(* IEC 61131-3 sources: guidance-for-physical-ai-production-designer-on-aws/source/plan2cell/examples/cell_2robot/plc/codesys/robots/robot1/GVL, 3 files *)

(* ---- GVL_DeviceParams.st ---- *)
(*
 * GVL_DeviceParams
 * PROFINET device identity parameters.
 * Device simulator R1 (robot1, station kuka-robi1), cell cell_2robot. Generated by bt2plc 0.1.0.
 *
 * These parameters configure how the CODESYS PROFINET Device presents itself
 * on the network. They MUST match what the Siemens PLC expects (from the GSDML).
 *
 * In CODESYS, these are typically set via:
 *   1. The "PROFINET Device IEC Objects" tab in the device editor
 *   2. Or programmatically by writing to the device parameter structure
 *
 * The CODESYS PROFINET Device stack reads these at startup and uses them
 * in DCP responses and during the PROFINET connection establishment.
 *
 * IMPORTANT: The default CODESYS values (VendorId=0x02CC, DeviceId=0x1017)
 * will NOT work with the Siemens PLC that expects KUKA (0x019B / 0x0301).
 * You MUST override them.
 *)

{attribute 'qualified_only'}
VAR_GLOBAL CONSTANT
    (* === KUKA VKRCnexxt Device Identity === *)
    (* These values come from GSDML-V2.25-KUKA-Roboter-GmbH-VKR C4-Device-V1.0 *)

    VENDOR_ID           : UINT        := 16#019B;                 (* KUKA Roboter GmbH *)
    DEVICE_ID           : UINT        := 16#0301;                 (* VKR C4 Device *)
    STATION_TYPE        : STRING(240) := 'KUKA VKR C4';           (* Station type string *)
    DEVICE_TYPE         : STRING(28)  := 'KUKA VKR C4';           (* Device type string *)
    ORDER_ID            : STRING(20)  := 'KUKA VKRC nexxt';       (* Order number *)
    HW_REVISION         : UINT        := 1;                       (* Hardware revision *)
    SW_REV_PREFIX       : USINT       := 16#56;                   (* 'V' in ASCII *)
    SW_REV_MAJOR        : UINT        := 8;                       (* V8.x *)
    SW_REV_MINOR        : UINT        := 2;                       (* x.2 *)
    SW_REV_PATCH        : UINT        := 0;                       (* x.x.0 *)

    (* === Module Identification Numbers (from GSDML) === *)
    MODULE_IDENT_DAP    : DWORD       := DWORD#16#00000301;       (* DAP - Slot 0 *)
    MODULE_IDENT_FDIO64 : DWORD       := DWORD#16#0000008F;       (* PROFIsafe - Slot 1 *)
    MODULE_IDENT_DIO256 : DWORD       := DWORD#16#00001000;       (* VASS telegram - Slot 2 *)
    SUBMODULE_IDENT     : DWORD       := DWORD#16#00000001;       (* Submodule ident (all slots) *)

    (* === PROFIsafe Parameters (Slot 1) === *)
    (* These must match the F-parameter record in the PLC safety configuration *)
    F_SIL_LEVEL         : UINT        := 3;                       (* SIL 3 *)
    F_CRC_LENGTH        : UINT        := 3;                       (* 3-byte CRC *)
    F_WD_TIME_DEFAULT   : UINT        := 500;                     (* Watchdog 500ms *)
    F_BLOCK_ID          : UINT        := 0;                       (* Block ID *)
    F_PAR_CRC_DEFAULT   : UINT        := 16#FF59;                 (* Default F_Par_CRC = 65369 *)
END_VAR

(* ---- GVL_IO.st ---- *)
(*
 * GVL_IO
 * Global variable list for the PROFINET device I/O mapping.
 * Device simulator R1 (robot1, station kuka-robi1), cell cell_2robot. Generated by bt2plc 0.1.0.
 *
 * These variables are mapped to the PROFINET device modules via the I/O Mapping tab.
 * Do NOT use AT addresses - the mapping is done in the device configuration.
 * Only PLC_PRG accesses this GVL: it copies the commands into local images and writes
 * the robot status back as a whole array / as scalars (the FBs never touch GVL_IO).
 *
 * Module mapping (set in I/O Mapping tab of each module):
 *   SafeIO_FDIO64 (Slot 1):
 *     "8 safe digital inputs" channels  -> GVL_IO.bySafeIn0..bySafeIn7
 *     "8 safe digital outputs" channels -> GVL_IO.bySafeOut0..bySafeOut7
 *
 *   VASS_DIO256 (Slot 2):
 *     Input channel  -> GVL_IO.aVassInputData
 *     Output channel -> GVL_IO.aVassOutputData
 *)

{attribute 'qualified_only'}
VAR_GLOBAL
    (* ========================================================================
       SLOT 1 - PROFIsafe FDIO64 Module
       8 individual USINT/BYTE channels per direction
       Map each one to the corresponding "8 safe digital inputs/outputs" row
       ======================================================================== *)

    (* Safe Inputs: Robot -> PLC (mapped to "8 safe digital inputs" channels) *)
    bySafeIn0       : BYTE;     (* Safe input byte 0: Drive status *)
    bySafeIn1       : BYTE;     (* Safe input byte 1: Gate/protection *)
    bySafeIn2       : BYTE;     (* Safe input byte 2: STO/SS1/SS2/SOS/SLS *)
    bySafeIn3       : BYTE;     (* Safe input byte 3: User *)
    bySafeIn4       : BYTE;     (* Safe input byte 4: User *)
    bySafeIn5       : BYTE;     (* Safe input byte 5: User *)
    bySafeIn6       : BYTE;     (* Safe input byte 6: User *)
    bySafeIn7       : BYTE;     (* Safe input byte 7: User *)

    (* Safe Outputs: PLC -> Robot (mapped to "8 safe digital outputs" channels) *)
    bySafeOut0      : BYTE;     (* Safe output byte 0: Drive enable, E-Stop, SS1/SS2 *)
    bySafeOut1      : BYTE;     (* Safe output byte 1: Zone enables *)
    bySafeOut2      : BYTE;     (* Safe output byte 2: User *)
    bySafeOut3      : BYTE;     (* Safe output byte 3: User *)
    bySafeOut4      : BYTE;     (* Safe output byte 4: User *)
    bySafeOut5      : BYTE;     (* Safe output byte 5: User *)
    bySafeOut6      : BYTE;     (* Safe output byte 6: User *)
    bySafeOut7      : BYTE;     (* Safe output byte 7: User *)

    (* ========================================================================
       SLOT 2 - DIO256 VASS Telegram
       32 bytes per direction as arrays
       ======================================================================== *)

    (* VASS Inputs: Robot -> PLC (32 bytes) *)
    aVassInputData      : ARRAY[0..31] OF BYTE;

    (* VASS Outputs: PLC -> Robot (32 bytes) *)
    aVassOutputData     : ARRAY[0..31] OF BYTE;
END_VAR

(* ---- GVL_Program.st ---- *)
(*
 * GVL_Program - generated by bt2plc 0.1.0 - DO NOT EDIT
 * Robot program of robot1 (R1) for plan bt_1791274820_cell_2robot (cell cell_2robot)
 * Angles in degrees (KUKA A1..A6 after joint sign/offset), times in seconds from op start.
 *)
{attribute 'qualified_only'}
VAR_GLOBAL CONSTANT
    (* ========================================================================
       IDENTITY / PROTOCOL
       ======================================================================== *)
    ROBOT_TAG               : STRING(16) := 'R1';
    ROBOT_NS                : STRING(32) := 'robot1';
    ROBOT_INDEX             : WORD := WORD#1;
    PLAN_ID                 : WORD := WORD#16#A312;             (* must match the head PLC *)
    PROD_FOLGE              : WORD := WORD#11;
    HOME_FOLGE              : WORD := WORD#125;
    JOB_NUMBER_BYTE         : BOOL := FALSE;
    STEP_BYTE               : INT := 4;
    REQ_BYTE                : INT := 28;
    GRANT_BYTE              : INT := 12;
    PLAN_ID_BYTE            : INT := 4;
    R_TASK_S                : REAL := 0.0200;                   (* device MainTask interval *)
    R_HOME_S                : REAL := 7.0000;                   (* blind home duration *)
    R_AT_HOME_TOL_DEG       : REAL := 0.5000;
    R_START_TOL_DEG         : REAL := 1.0000;
    ERR_UNKNOWN_FOLGE       : WORD := WORD#16#0101;
    ERR_PLAN_MISMATCH       : WORD := WORD#16#0103;
    WARN_START_DEVIATION    : WORD := WORD#16#0201;

    (* ========================================================================
       PROGRAM
       ======================================================================== *)
    N_OPS                   : INT := 2;
    N_WP                    : INT := 27;
    arHomeDeg               : ARRAY[1..6] OF REAL := [0.0000, -90.0000, 90.0000, 0.0000, 0.0000, 0.0000];
    aOps                    : ARRAY[1..2] OF ST_OpDef := [
        (sName := 'STAGE_R1', nFirstWp := 1, nLastWp := 14, dwZoneMask := DWORD#16#00000000, tDelay := T#0MS, tHold := T#500MS, rDelay_s := 0.0000, rHold_s := 0.5000, rVelScale := 1.0000, bBlindHome := FALSE),    (* #1 STAGE_R1 (move) *)
        (sName := 'HOME', nFirstWp := 15, nLastWp := 27, dwZoneMask := DWORD#16#00000000, tDelay := T#0MS, tHold := T#0MS, rDelay_s := 0.0000, rHold_s := 0.0000, rVelScale := 1.0000, bBlindHome := FALSE)    (* #2 HOME (home) *)
    ];
    aWp                     : ARRAY[1..27] OF ST_Waypoint := [
        (* op 1 STAGE_R1 - traj_robot1_STAGE_R1 *)
        (rT := 0.0000, rA1 := 0.0000, rA2 := -90.0000, rA3 := 90.0000, rA4 := 0.0000, rA5 := 0.0000, rA6 := 0.0000),
        (rT := 0.2767, rA1 := 0.1421, rA2 := -89.0006, rA3 := 89.9771, rA4 := 0.0000, rA5 := 0.0000, rA6 := 0.0000),
        (rT := 0.5530, rA1 := 0.5354, rA2 := -86.2310, rA3 := 89.9133, rA4 := 0.0000, rA5 := 0.0000, rA6 := 0.0000),
        (rT := 0.8297, rA1 := 1.1310, rA2 := -82.0342, rA3 := 89.8161, rA4 := 0.0000, rA5 := 0.0000, rA6 := 0.0000),
        (rT := 1.1063, rA1 := 1.8795, rA2 := -76.7531, rA3 := 89.6931, rA4 := 0.0000, rA5 := 0.0000, rA6 := 0.0000),
        (rT := 1.3830, rA1 := 2.7319, rA2 := -70.7305, rA3 := 89.5515, rA4 := 0.0000, rA5 := 0.0000, rA6 := 0.0000),
        (rT := 1.6593, rA1 := 3.6388, rA2 := -64.3095, rA3 := 89.3990, rA4 := 0.0000, rA5 := 0.0000, rA6 := 0.0000),
        (rT := 1.9360, rA1 := 4.5513, rA2 := -57.8329, rA3 := 89.2429, rA4 := 0.0000, rA5 := 0.0000, rA6 := 0.0000),
        (rT := 2.2127, rA1 := 5.4200, rA2 := -51.6436, rA3 := 89.0908, rA4 := 0.0000, rA5 := 0.0000, rA6 := 0.0000),
        (rT := 2.4893, rA1 := 6.1959, rA2 := -46.0847, rA3 := 88.9501, rA4 := 0.0000, rA5 := 0.0000, rA6 := 0.0000),
        (rT := 2.7657, rA1 := 6.8297, rA2 := -41.4990, rA3 := 88.8283, rA4 := 0.0000, rA5 := 0.0000, rA6 := 0.0000),
        (rT := 3.0423, rA1 := 7.2722, rA2 := -38.2294, rA3 := 88.7329, rA4 := 0.0000, rA5 := 0.0000, rA6 := 0.0000),
        (rT := 3.1357, rA1 := 7.7267, rA2 := -33.2119, rA3 := 88.3788, rA4 := 0.0000, rA5 := 0.0000, rA6 := 0.0000),
        (rT := 3.2287, rA1 := 7.2722, rA2 := -35.0616, rA3 := 88.2443, rA4 := 0.0000, rA5 := 0.0000, rA6 := 0.0000),
        (* op 2 HOME - traj_robot1_n3 *)
        (rT := 0.0000, rA1 := 7.2722, rA2 := -35.0616, rA3 := 88.2443, rA4 := 0.0000, rA5 := 0.0000, rA6 := 0.0000),
        (rT := 0.2015, rA1 := 7.1292, rA2 := -36.1426, rA3 := 88.2788, rA4 := 0.0000, rA5 := 0.0000, rA6 := 0.0000),
        (rT := 0.4032, rA1 := 6.7336, rA2 := -39.1311, rA3 := 88.3743, rA4 := 0.0000, rA5 := 0.0000, rA6 := 0.0000),
        (rT := 0.6048, rA1 := 6.1360, rA2 := -43.6457, rA3 := 88.5186, rA4 := 0.0000, rA5 := 0.0000, rA6 := 0.0000),
        (rT := 0.8065, rA1 := 5.3868, rA2 := -49.3049, rA3 := 88.6995, rA4 := 0.0000, rA5 := 0.0000, rA6 := 0.0000),
        (rT := 1.0080, rA1 := 4.5367, rA2 := -55.7271, rA3 := 88.9047, rA4 := 0.0000, rA5 := 0.0000, rA6 := 0.0000),
        (rT := 1.2097, rA1 := 3.6361, rA2 := -62.5308, rA3 := 89.1221, rA4 := 0.0000, rA5 := 0.0000, rA6 := 0.0000),
        (rT := 1.4112, rA1 := 2.7355, rA2 := -69.3345, rA3 := 89.3396, rA4 := 0.0000, rA5 := 0.0000, rA6 := 0.0000),
        (rT := 1.6127, rA1 := 1.8854, rA2 := -75.7567, rA3 := 89.5448, rA4 := 0.0000, rA5 := 0.0000, rA6 := 0.0000),
        (rT := 1.8145, rA1 := 1.1363, rA2 := -81.4159, rA3 := 89.7257, rA4 := 0.0000, rA5 := 0.0000, rA6 := 0.0000),
        (rT := 2.0160, rA1 := 0.5387, rA2 := -85.9305, rA3 := 89.8699, rA4 := 0.0000, rA5 := 0.0000, rA6 := 0.0000),
        (rT := 2.2177, rA1 := 0.1431, rA2 := -88.9190, rA3 := 89.9655, rA4 := 0.0000, rA5 := 0.0000, rA6 := 0.0000),
        (rT := 2.4192, rA1 := 0.0000, rA2 := -90.0000, rA3 := 90.0000, rA4 := 0.0000, rA5 := 0.0000, rA6 := 0.0000)
    ];
END_VAR
